# EPICS autosave request: 1.5.0/debian-12/7.0.10/modules/ADCore-ee039d2/db/NDArrayBase_settings.req
$(P)$(R)DataType
$(P)$(R)ColorMode
$(P)$(R)ArrayCallbacks
$(P)$(R)NDAttributesFile
$(P)$(R)NDAttributesMacros
$(P)$(R)PoolPollStats.SCAN
$(P)$(R)NumPreAllocBuffers
$(P)$(R)WaitForPlugins
